{attribute 'qualified_only'}
{attribute 'strict'}
TYPE E_CIP_DashStage :
(
	eCIPStage_NotInUse:= 0,
	eCIPStage_NotAvalable,
	eCIPStage_ToBeDone,
	eCIPStage_Active,
	eCIPStage_Done
);
END_TYPE

(* stored: Version 1.1.0.1, ProductVersion 3.1.4024.13
   DUT E_CIP_DashStage: Id {64f370dd-0aec-4a35-8d8d-41811d342d78} *)
